{attribute 'qualified_only'}
{attribute 'strict'}
TYPE E_TestStatus :
(
	Unknown := 0,
	Running,
	Passed,
	Failed,
	Aborted
);
END_TYPE

(* stored: Version 1.1.0.1, ProductVersion 3.1.4024.15
   DUT E_TestStatus: Id {338ac160-7013-4881-b326-13bd949cceb7} *)
